TYPE ST_ModeManagerActions :
STRUCT
    consumeResetReq : BOOL;
    clearModeFlags : BOOL;
    incrementResetAckCounter : BOOL;
    incrementWatchdogTripCounter : BOOL;
END_STRUCT
END_TYPE

(* stored: Version 1.1.0.1
   DUT ST_ModeManagerActions: Id {1E5573CE-A3E2-45EA-8707-49B3B9A7061E} *)
